(* IEC 61131-3 sources: s7-to-codesys/tests/POUs/ScenariosLang/FB_PumpInterlockLad_ScenarioTest, 6 files *)

(* ---- FB_PumpInterlockLad_ScenarioTest.decl.st ---- *)
// AUTO-GENERATED — не редактировать: s7conv gen-tests, сценарии scenarios/lang/FB_PumpInterlockLad.csv
// Правка — в CSV (scenarios/README.md), затем python -m s7conv build-corpus.
// Назначение: тесты поведения сконвертированного FB_PumpInterlockLad по сценариям CSV (сценариев: 5, строк: 25):
//             один метод-тест на сценарий, строки — по порядку с моделируемым временем GVL_S7Clock.
//             Ожидаемые значения — из CSV (эталонные модели по описанию логики блока), не из
//             результата конвертации.
// Автор:      s7conv 0.1.0 (сгенерировано)
// Версия:     не указана
// Документ:   scenarios/README.md, docs/methodology.md, раздел «Проверка поведения»
FUNCTION_BLOCK FB_PumpInterlockLad_ScenarioTest EXTENDS coUnit.FB_TestSuite
VAR
    fbAutoRunAndCount : FB_PumpInterlockLad;  // свой экземпляр на сценарий
    xAutoRunAndCountDone : BOOL;  // сценарий выполнен (выполняется один раз)
    fbLowLevelTripAndAck : FB_PumpInterlockLad;  // свой экземпляр на сценарий
    xLowLevelTripAndAckDone : BOOL;  // сценарий выполнен (выполняется один раз)
    fbHighPressure : FB_PumpInterlockLad;  // свой экземпляр на сценарий
    xHighPressureDone : BOOL;  // сценарий выполнен (выполняется один раз)
    fbMaintenanceJump : FB_PumpInterlockLad;  // свой экземпляр на сценарий
    xMaintenanceJumpDone : BOOL;  // сценарий выполнен (выполняется один раз)
    fbSetpointClamp : FB_PumpInterlockLad;  // свой экземпляр на сценарий
    xSetpointClampDone : BOOL;  // сценарий выполнен (выполняется один раз)
END_VAR

(* ---- AutoRunAndCount.method.impl.st ---- *)
// AUTO-GENERATED — не редактировать: scenarios/lang/FB_PumpInterlockLad.csv, сценарий AutoRunAndCount
coUnit.TEST('AutoRunAndCount');
IF NOT xAutoRunAndCountDone THEN
    xAutoRunAndCountDone := TRUE;
    GVL_S7Clock.xSimulation := TRUE;

    // #1, t = 0 мс — покой: уставка 0
    GVL_S7Clock.tSimNow := T#0MS;
    fbAutoRunAndCount.xAutoReq := FALSE;
    fbAutoRunAndCount.iLevel_cm := 120;
    fbAutoRunAndCount.iLevelMin_cm := 50;
    fbAutoRunAndCount.iPressure_kPa := 400;
    fbAutoRunAndCount.iPressureMax_kPa := 600;
    fbAutoRunAndCount.xAck := FALSE;
    fbAutoRunAndCount.xMaint := FALSE;
    fbAutoRunAndCount();
    AssertEquals_BOOL(Expected := FALSE, Actual := fbAutoRunAndCount.xPumpOn, Message := 'AutoRunAndCount#1 xPumpOn');
    AssertEquals_BOOL(Expected := FALSE,
                      Actual := fbAutoRunAndCount.xLowLevel,
                      Message := 'AutoRunAndCount#1 xLowLevel');
    AssertEquals_BOOL(Expected := FALSE,
                      Actual := fbAutoRunAndCount.xHighPress,
                      Message := 'AutoRunAndCount#1 xHighPress');
    AssertEquals_BOOL(Expected := FALSE, Actual := fbAutoRunAndCount.xAlarm, Message := 'AutoRunAndCount#1 xAlarm');
    AssertEquals_INT(Expected := 0, Actual := fbAutoRunAndCount.iRunCount, Message := 'AutoRunAndCount#1 iRunCount');
    AssertEquals_BOOL(Expected := FALSE, Actual := fbAutoRunAndCount.xCountOk, Message := 'AutoRunAndCount#1 xCountOk');
    AssertEquals_INT(Expected := 0,
                     Actual := fbAutoRunAndCount.iSetpoint_pct,
                     Message := 'AutoRunAndCount#1 iSetpoint_pct');
    AssertEquals_BOOL(Expected := FALSE, Actual := fbAutoRunAndCount.xChainOk, Message := 'AutoRunAndCount#1 xChainOk');
    AssertEquals_BOOL(Expected := FALSE, Actual := fbAutoRunAndCount.xRunMem, Message := 'AutoRunAndCount#1 xRunMem');

    // #2, t = 100 мс — включение №1: ENO = 1, уставка 120 → 100 → 90 → 80
    GVL_S7Clock.tSimNow := T#100MS;
    fbAutoRunAndCount.xAutoReq := TRUE;
    fbAutoRunAndCount();
    AssertEquals_BOOL(Expected := TRUE, Actual := fbAutoRunAndCount.xPumpOn, Message := 'AutoRunAndCount#2 xPumpOn');
    AssertEquals_BOOL(Expected := FALSE,
                      Actual := fbAutoRunAndCount.xLowLevel,
                      Message := 'AutoRunAndCount#2 xLowLevel');
    AssertEquals_BOOL(Expected := FALSE,
                      Actual := fbAutoRunAndCount.xHighPress,
                      Message := 'AutoRunAndCount#2 xHighPress');
    AssertEquals_BOOL(Expected := FALSE, Actual := fbAutoRunAndCount.xAlarm, Message := 'AutoRunAndCount#2 xAlarm');
    AssertEquals_INT(Expected := 1, Actual := fbAutoRunAndCount.iRunCount, Message := 'AutoRunAndCount#2 iRunCount');
    AssertEquals_BOOL(Expected := TRUE, Actual := fbAutoRunAndCount.xCountOk, Message := 'AutoRunAndCount#2 xCountOk');
    AssertEquals_INT(Expected := 80,
                     Actual := fbAutoRunAndCount.iSetpoint_pct,
                     Message := 'AutoRunAndCount#2 iSetpoint_pct');
    AssertEquals_BOOL(Expected := TRUE, Actual := fbAutoRunAndCount.xChainOk, Message := 'AutoRunAndCount#2 xChainOk');
    AssertEquals_BOOL(Expected := TRUE, Actual := fbAutoRunAndCount.xRunMem, Message := 'AutoRunAndCount#2 xRunMem');

    // #3, t = 200 мс — работает: фронта нет, ENO = 0
    GVL_S7Clock.tSimNow := T#200MS;
    fbAutoRunAndCount();
    AssertEquals_BOOL(Expected := TRUE, Actual := fbAutoRunAndCount.xPumpOn, Message := 'AutoRunAndCount#3 xPumpOn');
    AssertEquals_BOOL(Expected := FALSE,
                      Actual := fbAutoRunAndCount.xLowLevel,
                      Message := 'AutoRunAndCount#3 xLowLevel');
    AssertEquals_BOOL(Expected := FALSE,
                      Actual := fbAutoRunAndCount.xHighPress,
                      Message := 'AutoRunAndCount#3 xHighPress');
    AssertEquals_BOOL(Expected := FALSE, Actual := fbAutoRunAndCount.xAlarm, Message := 'AutoRunAndCount#3 xAlarm');
    AssertEquals_INT(Expected := 1, Actual := fbAutoRunAndCount.iRunCount, Message := 'AutoRunAndCount#3 iRunCount');
    AssertEquals_BOOL(Expected := FALSE, Actual := fbAutoRunAndCount.xCountOk, Message := 'AutoRunAndCount#3 xCountOk');
    AssertEquals_INT(Expected := 80,
                     Actual := fbAutoRunAndCount.iSetpoint_pct,
                     Message := 'AutoRunAndCount#3 iSetpoint_pct');
    AssertEquals_BOOL(Expected := TRUE, Actual := fbAutoRunAndCount.xChainOk, Message := 'AutoRunAndCount#3 xChainOk');
    AssertEquals_BOOL(Expected := TRUE, Actual := fbAutoRunAndCount.xRunMem, Message := 'AutoRunAndCount#3 xRunMem');

    // #4, t = 300 мс — запрос снят: насос выключен, уставка 0 (MOVE)
    GVL_S7Clock.tSimNow := T#300MS;
    fbAutoRunAndCount.xAutoReq := FALSE;
    fbAutoRunAndCount();
    AssertEquals_BOOL(Expected := FALSE, Actual := fbAutoRunAndCount.xPumpOn, Message := 'AutoRunAndCount#4 xPumpOn');
    AssertEquals_BOOL(Expected := FALSE,
                      Actual := fbAutoRunAndCount.xLowLevel,
                      Message := 'AutoRunAndCount#4 xLowLevel');
    AssertEquals_BOOL(Expected := FALSE,
                      Actual := fbAutoRunAndCount.xHighPress,
                      Message := 'AutoRunAndCount#4 xHighPress');
    AssertEquals_BOOL(Expected := FALSE, Actual := fbAutoRunAndCount.xAlarm, Message := 'AutoRunAndCount#4 xAlarm');
    AssertEquals_INT(Expected := 1, Actual := fbAutoRunAndCount.iRunCount, Message := 'AutoRunAndCount#4 iRunCount');
    AssertEquals_BOOL(Expected := FALSE, Actual := fbAutoRunAndCount.xCountOk, Message := 'AutoRunAndCount#4 xCountOk');
    AssertEquals_INT(Expected := 0,
                     Actual := fbAutoRunAndCount.iSetpoint_pct,
                     Message := 'AutoRunAndCount#4 iSetpoint_pct');
    AssertEquals_BOOL(Expected := FALSE, Actual := fbAutoRunAndCount.xChainOk, Message := 'AutoRunAndCount#4 xChainOk');
    AssertEquals_BOOL(Expected := FALSE, Actual := fbAutoRunAndCount.xRunMem, Message := 'AutoRunAndCount#4 xRunMem');

    // #5, t = 400 мс — включение №2
    GVL_S7Clock.tSimNow := T#400MS;
    fbAutoRunAndCount.xAutoReq := TRUE;
    fbAutoRunAndCount();
    AssertEquals_BOOL(Expected := TRUE, Actual := fbAutoRunAndCount.xPumpOn, Message := 'AutoRunAndCount#5 xPumpOn');
    AssertEquals_BOOL(Expected := FALSE,
                      Actual := fbAutoRunAndCount.xLowLevel,
                      Message := 'AutoRunAndCount#5 xLowLevel');
    AssertEquals_BOOL(Expected := FALSE,
                      Actual := fbAutoRunAndCount.xHighPress,
                      Message := 'AutoRunAndCount#5 xHighPress');
    AssertEquals_BOOL(Expected := FALSE, Actual := fbAutoRunAndCount.xAlarm, Message := 'AutoRunAndCount#5 xAlarm');
    AssertEquals_INT(Expected := 2, Actual := fbAutoRunAndCount.iRunCount, Message := 'AutoRunAndCount#5 iRunCount');
    AssertEquals_BOOL(Expected := TRUE, Actual := fbAutoRunAndCount.xCountOk, Message := 'AutoRunAndCount#5 xCountOk');
    AssertEquals_INT(Expected := 80,
                     Actual := fbAutoRunAndCount.iSetpoint_pct,
                     Message := 'AutoRunAndCount#5 iSetpoint_pct');
    AssertEquals_BOOL(Expected := TRUE, Actual := fbAutoRunAndCount.xChainOk, Message := 'AutoRunAndCount#5 xChainOk');
    AssertEquals_BOOL(Expected := TRUE, Actual := fbAutoRunAndCount.xRunMem, Message := 'AutoRunAndCount#5 xRunMem');

    GVL_S7Clock.xSimulation := FALSE;
END_IF
coUnit.TEST_FINISHED();

(* ---- HighPressure.method.impl.st ---- *)
// AUTO-GENERATED — не редактировать: scenarios/lang/FB_PumpInterlockLad.csv, сценарий HighPressure
coUnit.TEST('HighPressure');
IF NOT xHighPressureDone THEN
    xHighPressureDone := TRUE;
    GVL_S7Clock.xSimulation := TRUE;

    // #1, t = 0 мс — включение №1
    GVL_S7Clock.tSimNow := T#0MS;
    fbHighPressure.xAutoReq := TRUE;
    fbHighPressure.iLevel_cm := 120;
    fbHighPressure.iLevelMin_cm := 50;
    fbHighPressure.iPressure_kPa := 400;
    fbHighPressure.iPressureMax_kPa := 600;
    fbHighPressure.xAck := FALSE;
    fbHighPressure.xMaint := FALSE;
    fbHighPressure();
    AssertEquals_BOOL(Expected := TRUE, Actual := fbHighPressure.xPumpOn, Message := 'HighPressure#1 xPumpOn');
    AssertEquals_BOOL(Expected := FALSE, Actual := fbHighPressure.xLowLevel, Message := 'HighPressure#1 xLowLevel');
    AssertEquals_BOOL(Expected := FALSE, Actual := fbHighPressure.xHighPress, Message := 'HighPressure#1 xHighPress');
    AssertEquals_BOOL(Expected := FALSE, Actual := fbHighPressure.xAlarm, Message := 'HighPressure#1 xAlarm');
    AssertEquals_INT(Expected := 1, Actual := fbHighPressure.iRunCount, Message := 'HighPressure#1 iRunCount');
    AssertEquals_BOOL(Expected := TRUE, Actual := fbHighPressure.xCountOk, Message := 'HighPressure#1 xCountOk');
    AssertEquals_INT(Expected := 80, Actual := fbHighPressure.iSetpoint_pct, Message := 'HighPressure#1 iSetpoint_pct');
    AssertEquals_BOOL(Expected := TRUE, Actual := fbHighPressure.xChainOk, Message := 'HighPressure#1 xChainOk');
    AssertEquals_BOOL(Expected := TRUE, Actual := fbHighPressure.xRunMem, Message := 'HighPressure#1 xRunMem');

    // #2, t = 100 мс — 650 > 600: авария, насос выключен
    GVL_S7Clock.tSimNow := T#100MS;
    fbHighPressure.iPressure_kPa := 650;
    fbHighPressure();
    AssertEquals_BOOL(Expected := FALSE, Actual := fbHighPressure.xPumpOn, Message := 'HighPressure#2 xPumpOn');
    AssertEquals_BOOL(Expected := FALSE, Actual := fbHighPressure.xLowLevel, Message := 'HighPressure#2 xLowLevel');
    AssertEquals_BOOL(Expected := TRUE, Actual := fbHighPressure.xHighPress, Message := 'HighPressure#2 xHighPress');
    AssertEquals_BOOL(Expected := TRUE, Actual := fbHighPressure.xAlarm, Message := 'HighPressure#2 xAlarm');
    AssertEquals_INT(Expected := 1, Actual := fbHighPressure.iRunCount, Message := 'HighPressure#2 iRunCount');
    AssertEquals_BOOL(Expected := FALSE, Actual := fbHighPressure.xCountOk, Message := 'HighPressure#2 xCountOk');
    AssertEquals_INT(Expected := 0, Actual := fbHighPressure.iSetpoint_pct, Message := 'HighPressure#2 iSetpoint_pct');
    AssertEquals_BOOL(Expected := FALSE, Actual := fbHighPressure.xChainOk, Message := 'HighPressure#2 xChainOk');
    AssertEquals_BOOL(Expected := FALSE, Actual := fbHighPressure.xRunMem, Message := 'HighPressure#2 xRunMem');

    // #3, t = 200 мс — 600 не больше 600: квитирование снимает, включение №2
    GVL_S7Clock.tSimNow := T#200MS;
    fbHighPressure.iPressure_kPa := 600;
    fbHighPressure.xAck := TRUE;
    fbHighPressure();
    AssertEquals_BOOL(Expected := TRUE, Actual := fbHighPressure.xPumpOn, Message := 'HighPressure#3 xPumpOn');
    AssertEquals_BOOL(Expected := FALSE, Actual := fbHighPressure.xLowLevel, Message := 'HighPressure#3 xLowLevel');
    AssertEquals_BOOL(Expected := FALSE, Actual := fbHighPressure.xHighPress, Message := 'HighPressure#3 xHighPress');
    AssertEquals_BOOL(Expected := FALSE, Actual := fbHighPressure.xAlarm, Message := 'HighPressure#3 xAlarm');
    AssertEquals_INT(Expected := 2, Actual := fbHighPressure.iRunCount, Message := 'HighPressure#3 iRunCount');
    AssertEquals_BOOL(Expected := TRUE, Actual := fbHighPressure.xCountOk, Message := 'HighPressure#3 xCountOk');
    AssertEquals_INT(Expected := 80, Actual := fbHighPressure.iSetpoint_pct, Message := 'HighPressure#3 iSetpoint_pct');
    AssertEquals_BOOL(Expected := TRUE, Actual := fbHighPressure.xChainOk, Message := 'HighPressure#3 xChainOk');
    AssertEquals_BOOL(Expected := TRUE, Actual := fbHighPressure.xRunMem, Message := 'HighPressure#3 xRunMem');

    // #4, t = 300 мс — работает
    GVL_S7Clock.tSimNow := T#300MS;
    fbHighPressure.xAck := FALSE;
    fbHighPressure();
    AssertEquals_BOOL(Expected := TRUE, Actual := fbHighPressure.xPumpOn, Message := 'HighPressure#4 xPumpOn');
    AssertEquals_BOOL(Expected := FALSE, Actual := fbHighPressure.xLowLevel, Message := 'HighPressure#4 xLowLevel');
    AssertEquals_BOOL(Expected := FALSE, Actual := fbHighPressure.xHighPress, Message := 'HighPressure#4 xHighPress');
    AssertEquals_BOOL(Expected := FALSE, Actual := fbHighPressure.xAlarm, Message := 'HighPressure#4 xAlarm');
    AssertEquals_INT(Expected := 2, Actual := fbHighPressure.iRunCount, Message := 'HighPressure#4 iRunCount');
    AssertEquals_BOOL(Expected := FALSE, Actual := fbHighPressure.xCountOk, Message := 'HighPressure#4 xCountOk');
    AssertEquals_INT(Expected := 80, Actual := fbHighPressure.iSetpoint_pct, Message := 'HighPressure#4 iSetpoint_pct');
    AssertEquals_BOOL(Expected := TRUE, Actual := fbHighPressure.xChainOk, Message := 'HighPressure#4 xChainOk');
    AssertEquals_BOOL(Expected := TRUE, Actual := fbHighPressure.xRunMem, Message := 'HighPressure#4 xRunMem');

    GVL_S7Clock.xSimulation := FALSE;
END_IF
coUnit.TEST_FINISHED();

(* ---- LowLevelTripAndAck.method.impl.st ---- *)
// AUTO-GENERATED — не редактировать: scenarios/lang/FB_PumpInterlockLad.csv, сценарий LowLevelTripAndAck
coUnit.TEST('LowLevelTripAndAck');
IF NOT xLowLevelTripAndAckDone THEN
    xLowLevelTripAndAckDone := TRUE;
    GVL_S7Clock.xSimulation := TRUE;

    // #1, t = 0 мс — включение №1
    GVL_S7Clock.tSimNow := T#0MS;
    fbLowLevelTripAndAck.xAutoReq := TRUE;
    fbLowLevelTripAndAck.iLevel_cm := 120;
    fbLowLevelTripAndAck.iLevelMin_cm := 50;
    fbLowLevelTripAndAck.iPressure_kPa := 400;
    fbLowLevelTripAndAck.iPressureMax_kPa := 600;
    fbLowLevelTripAndAck.xAck := FALSE;
    fbLowLevelTripAndAck.xMaint := FALSE;
    fbLowLevelTripAndAck();
    AssertEquals_BOOL(Expected := TRUE,
                      Actual := fbLowLevelTripAndAck.xPumpOn,
                      Message := 'LowLevelTripAndAck#1 xPumpOn');
    AssertEquals_BOOL(Expected := FALSE,
                      Actual := fbLowLevelTripAndAck.xLowLevel,
                      Message := 'LowLevelTripAndAck#1 xLowLevel');
    AssertEquals_BOOL(Expected := FALSE,
                      Actual := fbLowLevelTripAndAck.xHighPress,
                      Message := 'LowLevelTripAndAck#1 xHighPress');
    AssertEquals_BOOL(Expected := FALSE,
                      Actual := fbLowLevelTripAndAck.xAlarm,
                      Message := 'LowLevelTripAndAck#1 xAlarm');
    AssertEquals_INT(Expected := 1,
                     Actual := fbLowLevelTripAndAck.iRunCount,
                     Message := 'LowLevelTripAndAck#1 iRunCount');
    AssertEquals_BOOL(Expected := TRUE,
                      Actual := fbLowLevelTripAndAck.xCountOk,
                      Message := 'LowLevelTripAndAck#1 xCountOk');
    AssertEquals_INT(Expected := 80,
                     Actual := fbLowLevelTripAndAck.iSetpoint_pct,
                     Message := 'LowLevelTripAndAck#1 iSetpoint_pct');
    AssertEquals_BOOL(Expected := TRUE,
                      Actual := fbLowLevelTripAndAck.xChainOk,
                      Message := 'LowLevelTripAndAck#1 xChainOk');
    AssertEquals_BOOL(Expected := TRUE,
                      Actual := fbLowLevelTripAndAck.xRunMem,
                      Message := 'LowLevelTripAndAck#1 xRunMem');

    // #2, t = 100 мс — уровень 40 < 50: авария, насос выключен
    GVL_S7Clock.tSimNow := T#100MS;
    fbLowLevelTripAndAck.iLevel_cm := 40;
    fbLowLevelTripAndAck();
    AssertEquals_BOOL(Expected := FALSE,
                      Actual := fbLowLevelTripAndAck.xPumpOn,
                      Message := 'LowLevelTripAndAck#2 xPumpOn');
    AssertEquals_BOOL(Expected := TRUE,
                      Actual := fbLowLevelTripAndAck.xLowLevel,
                      Message := 'LowLevelTripAndAck#2 xLowLevel');
    AssertEquals_BOOL(Expected := FALSE,
                      Actual := fbLowLevelTripAndAck.xHighPress,
                      Message := 'LowLevelTripAndAck#2 xHighPress');
    AssertEquals_BOOL(Expected := TRUE,
                      Actual := fbLowLevelTripAndAck.xAlarm,
                      Message := 'LowLevelTripAndAck#2 xAlarm');
    AssertEquals_INT(Expected := 1,
                     Actual := fbLowLevelTripAndAck.iRunCount,
                     Message := 'LowLevelTripAndAck#2 iRunCount');
    AssertEquals_BOOL(Expected := FALSE,
                      Actual := fbLowLevelTripAndAck.xCountOk,
                      Message := 'LowLevelTripAndAck#2 xCountOk');
    AssertEquals_INT(Expected := 0,
                     Actual := fbLowLevelTripAndAck.iSetpoint_pct,
                     Message := 'LowLevelTripAndAck#2 iSetpoint_pct');
    AssertEquals_BOOL(Expected := FALSE,
                      Actual := fbLowLevelTripAndAck.xChainOk,
                      Message := 'LowLevelTripAndAck#2 xChainOk');
    AssertEquals_BOOL(Expected := FALSE,
                      Actual := fbLowLevelTripAndAck.xRunMem,
                      Message := 'LowLevelTripAndAck#2 xRunMem');

    // #3, t = 200 мс — уровень в норме: авария держится
    GVL_S7Clock.tSimNow := T#200MS;
    fbLowLevelTripAndAck.iLevel_cm := 60;
    fbLowLevelTripAndAck();
    AssertEquals_BOOL(Expected := FALSE,
                      Actual := fbLowLevelTripAndAck.xPumpOn,
                      Message := 'LowLevelTripAndAck#3 xPumpOn');
    AssertEquals_BOOL(Expected := FALSE,
                      Actual := fbLowLevelTripAndAck.xLowLevel,
                      Message := 'LowLevelTripAndAck#3 xLowLevel');
    AssertEquals_BOOL(Expected := FALSE,
                      Actual := fbLowLevelTripAndAck.xHighPress,
                      Message := 'LowLevelTripAndAck#3 xHighPress');
    AssertEquals_BOOL(Expected := TRUE,
                      Actual := fbLowLevelTripAndAck.xAlarm,
                      Message := 'LowLevelTripAndAck#3 xAlarm');
    AssertEquals_INT(Expected := 1,
                     Actual := fbLowLevelTripAndAck.iRunCount,
                     Message := 'LowLevelTripAndAck#3 iRunCount');
    AssertEquals_BOOL(Expected := FALSE,
                      Actual := fbLowLevelTripAndAck.xCountOk,
                      Message := 'LowLevelTripAndAck#3 xCountOk');
    AssertEquals_INT(Expected := 0,
                     Actual := fbLowLevelTripAndAck.iSetpoint_pct,
                     Message := 'LowLevelTripAndAck#3 iSetpoint_pct');
    AssertEquals_BOOL(Expected := FALSE,
                      Actual := fbLowLevelTripAndAck.xChainOk,
                      Message := 'LowLevelTripAndAck#3 xChainOk');
    AssertEquals_BOOL(Expected := FALSE,
                      Actual := fbLowLevelTripAndAck.xRunMem,
                      Message := 'LowLevelTripAndAck#3 xRunMem');

    // #4, t = 300 мс — квитирование при низком уровне: не снимается
    GVL_S7Clock.tSimNow := T#300MS;
    fbLowLevelTripAndAck.iLevel_cm := 45;
    fbLowLevelTripAndAck.xAck := TRUE;
    fbLowLevelTripAndAck();
    AssertEquals_BOOL(Expected := FALSE,
                      Actual := fbLowLevelTripAndAck.xPumpOn,
                      Message := 'LowLevelTripAndAck#4 xPumpOn');
    AssertEquals_BOOL(Expected := TRUE,
                      Actual := fbLowLevelTripAndAck.xLowLevel,
                      Message := 'LowLevelTripAndAck#4 xLowLevel');
    AssertEquals_BOOL(Expected := FALSE,
                      Actual := fbLowLevelTripAndAck.xHighPress,
                      Message := 'LowLevelTripAndAck#4 xHighPress');
    AssertEquals_BOOL(Expected := TRUE,
                      Actual := fbLowLevelTripAndAck.xAlarm,
                      Message := 'LowLevelTripAndAck#4 xAlarm');
    AssertEquals_INT(Expected := 1,
                     Actual := fbLowLevelTripAndAck.iRunCount,
                     Message := 'LowLevelTripAndAck#4 iRunCount');
    AssertEquals_BOOL(Expected := FALSE,
                      Actual := fbLowLevelTripAndAck.xCountOk,
                      Message := 'LowLevelTripAndAck#4 xCountOk');
    AssertEquals_INT(Expected := 0,
                     Actual := fbLowLevelTripAndAck.iSetpoint_pct,
                     Message := 'LowLevelTripAndAck#4 iSetpoint_pct');
    AssertEquals_BOOL(Expected := FALSE,
                      Actual := fbLowLevelTripAndAck.xChainOk,
                      Message := 'LowLevelTripAndAck#4 xChainOk');
    AssertEquals_BOOL(Expected := FALSE,
                      Actual := fbLowLevelTripAndAck.xRunMem,
                      Message := 'LowLevelTripAndAck#4 xRunMem');

    // #5, t = 400 мс — уровень в норме при нажатом квитировании: снята, включение №2
    GVL_S7Clock.tSimNow := T#400MS;
    fbLowLevelTripAndAck.iLevel_cm := 70;
    fbLowLevelTripAndAck();
    AssertEquals_BOOL(Expected := TRUE,
                      Actual := fbLowLevelTripAndAck.xPumpOn,
                      Message := 'LowLevelTripAndAck#5 xPumpOn');
    AssertEquals_BOOL(Expected := FALSE,
                      Actual := fbLowLevelTripAndAck.xLowLevel,
                      Message := 'LowLevelTripAndAck#5 xLowLevel');
    AssertEquals_BOOL(Expected := FALSE,
                      Actual := fbLowLevelTripAndAck.xHighPress,
                      Message := 'LowLevelTripAndAck#5 xHighPress');
    AssertEquals_BOOL(Expected := FALSE,
                      Actual := fbLowLevelTripAndAck.xAlarm,
                      Message := 'LowLevelTripAndAck#5 xAlarm');
    AssertEquals_INT(Expected := 2,
                     Actual := fbLowLevelTripAndAck.iRunCount,
                     Message := 'LowLevelTripAndAck#5 iRunCount');
    AssertEquals_BOOL(Expected := TRUE,
                      Actual := fbLowLevelTripAndAck.xCountOk,
                      Message := 'LowLevelTripAndAck#5 xCountOk');
    AssertEquals_INT(Expected := 70,
                     Actual := fbLowLevelTripAndAck.iSetpoint_pct,
                     Message := 'LowLevelTripAndAck#5 iSetpoint_pct');
    AssertEquals_BOOL(Expected := TRUE,
                      Actual := fbLowLevelTripAndAck.xChainOk,
                      Message := 'LowLevelTripAndAck#5 xChainOk');
    AssertEquals_BOOL(Expected := TRUE,
                      Actual := fbLowLevelTripAndAck.xRunMem,
                      Message := 'LowLevelTripAndAck#5 xRunMem');

    // #6, t = 500 мс — работает
    GVL_S7Clock.tSimNow := T#500MS;
    fbLowLevelTripAndAck.xAck := FALSE;
    fbLowLevelTripAndAck();
    AssertEquals_BOOL(Expected := TRUE,
                      Actual := fbLowLevelTripAndAck.xPumpOn,
                      Message := 'LowLevelTripAndAck#6 xPumpOn');
    AssertEquals_BOOL(Expected := FALSE,
                      Actual := fbLowLevelTripAndAck.xLowLevel,
                      Message := 'LowLevelTripAndAck#6 xLowLevel');
    AssertEquals_BOOL(Expected := FALSE,
                      Actual := fbLowLevelTripAndAck.xHighPress,
                      Message := 'LowLevelTripAndAck#6 xHighPress');
    AssertEquals_BOOL(Expected := FALSE,
                      Actual := fbLowLevelTripAndAck.xAlarm,
                      Message := 'LowLevelTripAndAck#6 xAlarm');
    AssertEquals_INT(Expected := 2,
                     Actual := fbLowLevelTripAndAck.iRunCount,
                     Message := 'LowLevelTripAndAck#6 iRunCount');
    AssertEquals_BOOL(Expected := FALSE,
                      Actual := fbLowLevelTripAndAck.xCountOk,
                      Message := 'LowLevelTripAndAck#6 xCountOk');
    AssertEquals_INT(Expected := 70,
                     Actual := fbLowLevelTripAndAck.iSetpoint_pct,
                     Message := 'LowLevelTripAndAck#6 iSetpoint_pct');
    AssertEquals_BOOL(Expected := TRUE,
                      Actual := fbLowLevelTripAndAck.xChainOk,
                      Message := 'LowLevelTripAndAck#6 xChainOk');
    AssertEquals_BOOL(Expected := TRUE,
                      Actual := fbLowLevelTripAndAck.xRunMem,
                      Message := 'LowLevelTripAndAck#6 xRunMem');

    GVL_S7Clock.xSimulation := FALSE;
END_IF
coUnit.TEST_FINISHED();

(* ---- MaintenanceJump.method.impl.st ---- *)
// AUTO-GENERATED — не редактировать: scenarios/lang/FB_PumpInterlockLad.csv, сценарий MaintenanceJump
coUnit.TEST('MaintenanceJump');
IF NOT xMaintenanceJumpDone THEN
    xMaintenanceJumpDone := TRUE;
    GVL_S7Clock.xSimulation := TRUE;

    // #1, t = 0 мс — включение №1, xCountOk = 1
    GVL_S7Clock.tSimNow := T#0MS;
    fbMaintenanceJump.xAutoReq := TRUE;
    fbMaintenanceJump.iLevel_cm := 120;
    fbMaintenanceJump.iLevelMin_cm := 50;
    fbMaintenanceJump.iPressure_kPa := 400;
    fbMaintenanceJump.iPressureMax_kPa := 600;
    fbMaintenanceJump.xAck := FALSE;
    fbMaintenanceJump.xMaint := FALSE;
    fbMaintenanceJump();
    AssertEquals_BOOL(Expected := TRUE, Actual := fbMaintenanceJump.xPumpOn, Message := 'MaintenanceJump#1 xPumpOn');
    AssertEquals_BOOL(Expected := FALSE,
                      Actual := fbMaintenanceJump.xLowLevel,
                      Message := 'MaintenanceJump#1 xLowLevel');
    AssertEquals_BOOL(Expected := FALSE,
                      Actual := fbMaintenanceJump.xHighPress,
                      Message := 'MaintenanceJump#1 xHighPress');
    AssertEquals_BOOL(Expected := FALSE, Actual := fbMaintenanceJump.xAlarm, Message := 'MaintenanceJump#1 xAlarm');
    AssertEquals_INT(Expected := 1, Actual := fbMaintenanceJump.iRunCount, Message := 'MaintenanceJump#1 iRunCount');
    AssertEquals_BOOL(Expected := TRUE, Actual := fbMaintenanceJump.xCountOk, Message := 'MaintenanceJump#1 xCountOk');
    AssertEquals_INT(Expected := 80,
                     Actual := fbMaintenanceJump.iSetpoint_pct,
                     Message := 'MaintenanceJump#1 iSetpoint_pct');
    AssertEquals_BOOL(Expected := TRUE, Actual := fbMaintenanceJump.xChainOk, Message := 'MaintenanceJump#1 xChainOk');
    AssertEquals_BOOL(Expected := TRUE, Actual := fbMaintenanceJump.xRunMem, Message := 'MaintenanceJump#1 xRunMem');

    // #2, t = 100 мс — обслуживание: насос выключен; xCountOk и xRunMem сохраняют значения
    GVL_S7Clock.tSimNow := T#100MS;
    fbMaintenanceJump.xMaint := TRUE;
    fbMaintenanceJump();
    AssertEquals_BOOL(Expected := FALSE, Actual := fbMaintenanceJump.xPumpOn, Message := 'MaintenanceJump#2 xPumpOn');
    AssertEquals_BOOL(Expected := FALSE,
                      Actual := fbMaintenanceJump.xLowLevel,
                      Message := 'MaintenanceJump#2 xLowLevel');
    AssertEquals_BOOL(Expected := FALSE,
                      Actual := fbMaintenanceJump.xHighPress,
                      Message := 'MaintenanceJump#2 xHighPress');
    AssertEquals_BOOL(Expected := FALSE, Actual := fbMaintenanceJump.xAlarm, Message := 'MaintenanceJump#2 xAlarm');
    AssertEquals_INT(Expected := 1, Actual := fbMaintenanceJump.iRunCount, Message := 'MaintenanceJump#2 iRunCount');
    AssertEquals_BOOL(Expected := TRUE, Actual := fbMaintenanceJump.xCountOk, Message := 'MaintenanceJump#2 xCountOk');
    AssertEquals_INT(Expected := 0,
                     Actual := fbMaintenanceJump.iSetpoint_pct,
                     Message := 'MaintenanceJump#2 iSetpoint_pct');
    AssertEquals_BOOL(Expected := FALSE, Actual := fbMaintenanceJump.xChainOk, Message := 'MaintenanceJump#2 xChainOk');
    AssertEquals_BOOL(Expected := TRUE, Actual := fbMaintenanceJump.xRunMem, Message := 'MaintenanceJump#2 xRunMem');

    // #3, t = 200 мс — обслуживание держится
    GVL_S7Clock.tSimNow := T#200MS;
    fbMaintenanceJump();
    AssertEquals_BOOL(Expected := FALSE, Actual := fbMaintenanceJump.xPumpOn, Message := 'MaintenanceJump#3 xPumpOn');
    AssertEquals_BOOL(Expected := FALSE,
                      Actual := fbMaintenanceJump.xLowLevel,
                      Message := 'MaintenanceJump#3 xLowLevel');
    AssertEquals_BOOL(Expected := FALSE,
                      Actual := fbMaintenanceJump.xHighPress,
                      Message := 'MaintenanceJump#3 xHighPress');
    AssertEquals_BOOL(Expected := FALSE, Actual := fbMaintenanceJump.xAlarm, Message := 'MaintenanceJump#3 xAlarm');
    AssertEquals_INT(Expected := 1, Actual := fbMaintenanceJump.iRunCount, Message := 'MaintenanceJump#3 iRunCount');
    AssertEquals_BOOL(Expected := TRUE, Actual := fbMaintenanceJump.xCountOk, Message := 'MaintenanceJump#3 xCountOk');
    AssertEquals_INT(Expected := 0,
                     Actual := fbMaintenanceJump.iSetpoint_pct,
                     Message := 'MaintenanceJump#3 iSetpoint_pct');
    AssertEquals_BOOL(Expected := FALSE, Actual := fbMaintenanceJump.xChainOk, Message := 'MaintenanceJump#3 xChainOk');
    AssertEquals_BOOL(Expected := TRUE, Actual := fbMaintenanceJump.xRunMem, Message := 'MaintenanceJump#3 xRunMem');

    // #4, t = 300 мс — выход из обслуживания: насос включён, фронта нет — бит памяти остался 1
    GVL_S7Clock.tSimNow := T#300MS;
    fbMaintenanceJump.xMaint := FALSE;
    fbMaintenanceJump();
    AssertEquals_BOOL(Expected := TRUE, Actual := fbMaintenanceJump.xPumpOn, Message := 'MaintenanceJump#4 xPumpOn');
    AssertEquals_BOOL(Expected := FALSE,
                      Actual := fbMaintenanceJump.xLowLevel,
                      Message := 'MaintenanceJump#4 xLowLevel');
    AssertEquals_BOOL(Expected := FALSE,
                      Actual := fbMaintenanceJump.xHighPress,
                      Message := 'MaintenanceJump#4 xHighPress');
    AssertEquals_BOOL(Expected := FALSE, Actual := fbMaintenanceJump.xAlarm, Message := 'MaintenanceJump#4 xAlarm');
    AssertEquals_INT(Expected := 1, Actual := fbMaintenanceJump.iRunCount, Message := 'MaintenanceJump#4 iRunCount');
    AssertEquals_BOOL(Expected := FALSE, Actual := fbMaintenanceJump.xCountOk, Message := 'MaintenanceJump#4 xCountOk');
    AssertEquals_INT(Expected := 80,
                     Actual := fbMaintenanceJump.iSetpoint_pct,
                     Message := 'MaintenanceJump#4 iSetpoint_pct');
    AssertEquals_BOOL(Expected := TRUE, Actual := fbMaintenanceJump.xChainOk, Message := 'MaintenanceJump#4 xChainOk');
    AssertEquals_BOOL(Expected := TRUE, Actual := fbMaintenanceJump.xRunMem, Message := 'MaintenanceJump#4 xRunMem');

    // #5, t = 400 мс — запрос снят
    GVL_S7Clock.tSimNow := T#400MS;
    fbMaintenanceJump.xAutoReq := FALSE;
    fbMaintenanceJump();
    AssertEquals_BOOL(Expected := FALSE, Actual := fbMaintenanceJump.xPumpOn, Message := 'MaintenanceJump#5 xPumpOn');
    AssertEquals_BOOL(Expected := FALSE,
                      Actual := fbMaintenanceJump.xLowLevel,
                      Message := 'MaintenanceJump#5 xLowLevel');
    AssertEquals_BOOL(Expected := FALSE,
                      Actual := fbMaintenanceJump.xHighPress,
                      Message := 'MaintenanceJump#5 xHighPress');
    AssertEquals_BOOL(Expected := FALSE, Actual := fbMaintenanceJump.xAlarm, Message := 'MaintenanceJump#5 xAlarm');
    AssertEquals_INT(Expected := 1, Actual := fbMaintenanceJump.iRunCount, Message := 'MaintenanceJump#5 iRunCount');
    AssertEquals_BOOL(Expected := FALSE, Actual := fbMaintenanceJump.xCountOk, Message := 'MaintenanceJump#5 xCountOk');
    AssertEquals_INT(Expected := 0,
                     Actual := fbMaintenanceJump.iSetpoint_pct,
                     Message := 'MaintenanceJump#5 iSetpoint_pct');
    AssertEquals_BOOL(Expected := FALSE, Actual := fbMaintenanceJump.xChainOk, Message := 'MaintenanceJump#5 xChainOk');
    AssertEquals_BOOL(Expected := FALSE, Actual := fbMaintenanceJump.xRunMem, Message := 'MaintenanceJump#5 xRunMem');

    // #6, t = 500 мс — включение №2
    GVL_S7Clock.tSimNow := T#500MS;
    fbMaintenanceJump.xAutoReq := TRUE;
    fbMaintenanceJump();
    AssertEquals_BOOL(Expected := TRUE, Actual := fbMaintenanceJump.xPumpOn, Message := 'MaintenanceJump#6 xPumpOn');
    AssertEquals_BOOL(Expected := FALSE,
                      Actual := fbMaintenanceJump.xLowLevel,
                      Message := 'MaintenanceJump#6 xLowLevel');
    AssertEquals_BOOL(Expected := FALSE,
                      Actual := fbMaintenanceJump.xHighPress,
                      Message := 'MaintenanceJump#6 xHighPress');
    AssertEquals_BOOL(Expected := FALSE, Actual := fbMaintenanceJump.xAlarm, Message := 'MaintenanceJump#6 xAlarm');
    AssertEquals_INT(Expected := 2, Actual := fbMaintenanceJump.iRunCount, Message := 'MaintenanceJump#6 iRunCount');
    AssertEquals_BOOL(Expected := TRUE, Actual := fbMaintenanceJump.xCountOk, Message := 'MaintenanceJump#6 xCountOk');
    AssertEquals_INT(Expected := 80,
                     Actual := fbMaintenanceJump.iSetpoint_pct,
                     Message := 'MaintenanceJump#6 iSetpoint_pct');
    AssertEquals_BOOL(Expected := TRUE, Actual := fbMaintenanceJump.xChainOk, Message := 'MaintenanceJump#6 xChainOk');
    AssertEquals_BOOL(Expected := TRUE, Actual := fbMaintenanceJump.xRunMem, Message := 'MaintenanceJump#6 xRunMem');

    GVL_S7Clock.xSimulation := FALSE;
END_IF
coUnit.TEST_FINISHED();

(* ---- SetpointClamp.method.impl.st ---- *)
// AUTO-GENERATED — не редактировать: scenarios/lang/FB_PumpInterlockLad.csv, сценарий SetpointClamp
coUnit.TEST('SetpointClamp');
IF NOT xSetpointClampDone THEN
    xSetpointClampDone := TRUE;
    GVL_S7Clock.xSimulation := TRUE;

    // #1, t = 0 мс — 55 → 55 → 55 → 55
    GVL_S7Clock.tSimNow := T#0MS;
    fbSetpointClamp.xAutoReq := TRUE;
    fbSetpointClamp.iLevel_cm := 55;
    fbSetpointClamp.iLevelMin_cm := 50;
    fbSetpointClamp.iPressure_kPa := 400;
    fbSetpointClamp.iPressureMax_kPa := 600;
    fbSetpointClamp.xAck := FALSE;
    fbSetpointClamp.xMaint := FALSE;
    fbSetpointClamp();
    AssertEquals_BOOL(Expected := TRUE, Actual := fbSetpointClamp.xPumpOn, Message := 'SetpointClamp#1 xPumpOn');
    AssertEquals_BOOL(Expected := FALSE, Actual := fbSetpointClamp.xLowLevel, Message := 'SetpointClamp#1 xLowLevel');
    AssertEquals_BOOL(Expected := FALSE, Actual := fbSetpointClamp.xHighPress, Message := 'SetpointClamp#1 xHighPress');
    AssertEquals_BOOL(Expected := FALSE, Actual := fbSetpointClamp.xAlarm, Message := 'SetpointClamp#1 xAlarm');
    AssertEquals_INT(Expected := 1, Actual := fbSetpointClamp.iRunCount, Message := 'SetpointClamp#1 iRunCount');
    AssertEquals_BOOL(Expected := TRUE, Actual := fbSetpointClamp.xCountOk, Message := 'SetpointClamp#1 xCountOk');
    AssertEquals_INT(Expected := 55,
                     Actual := fbSetpointClamp.iSetpoint_pct,
                     Message := 'SetpointClamp#1 iSetpoint_pct');
    AssertEquals_BOOL(Expected := TRUE, Actual := fbSetpointClamp.xChainOk, Message := 'SetpointClamp#1 xChainOk');
    AssertEquals_BOOL(Expected := TRUE, Actual := fbSetpointClamp.xRunMem, Message := 'SetpointClamp#1 xRunMem');

    // #2, t = 100 мс — 95 → 95 → 90 → 80
    GVL_S7Clock.tSimNow := T#100MS;
    fbSetpointClamp.iLevel_cm := 95;
    fbSetpointClamp();
    AssertEquals_BOOL(Expected := TRUE, Actual := fbSetpointClamp.xPumpOn, Message := 'SetpointClamp#2 xPumpOn');
    AssertEquals_BOOL(Expected := FALSE, Actual := fbSetpointClamp.xLowLevel, Message := 'SetpointClamp#2 xLowLevel');
    AssertEquals_BOOL(Expected := FALSE, Actual := fbSetpointClamp.xHighPress, Message := 'SetpointClamp#2 xHighPress');
    AssertEquals_BOOL(Expected := FALSE, Actual := fbSetpointClamp.xAlarm, Message := 'SetpointClamp#2 xAlarm');
    AssertEquals_INT(Expected := 1, Actual := fbSetpointClamp.iRunCount, Message := 'SetpointClamp#2 iRunCount');
    AssertEquals_BOOL(Expected := FALSE, Actual := fbSetpointClamp.xCountOk, Message := 'SetpointClamp#2 xCountOk');
    AssertEquals_INT(Expected := 80,
                     Actual := fbSetpointClamp.iSetpoint_pct,
                     Message := 'SetpointClamp#2 iSetpoint_pct');
    AssertEquals_BOOL(Expected := TRUE, Actual := fbSetpointClamp.xChainOk, Message := 'SetpointClamp#2 xChainOk');
    AssertEquals_BOOL(Expected := TRUE, Actual := fbSetpointClamp.xRunMem, Message := 'SetpointClamp#2 xRunMem');

    // #3, t = 200 мс — 15 → 15 → 15 → 20
    GVL_S7Clock.tSimNow := T#200MS;
    fbSetpointClamp.iLevel_cm := 15;
    fbSetpointClamp.iLevelMin_cm := 10;
    fbSetpointClamp();
    AssertEquals_BOOL(Expected := TRUE, Actual := fbSetpointClamp.xPumpOn, Message := 'SetpointClamp#3 xPumpOn');
    AssertEquals_BOOL(Expected := FALSE, Actual := fbSetpointClamp.xLowLevel, Message := 'SetpointClamp#3 xLowLevel');
    AssertEquals_BOOL(Expected := FALSE, Actual := fbSetpointClamp.xHighPress, Message := 'SetpointClamp#3 xHighPress');
    AssertEquals_BOOL(Expected := FALSE, Actual := fbSetpointClamp.xAlarm, Message := 'SetpointClamp#3 xAlarm');
    AssertEquals_INT(Expected := 1, Actual := fbSetpointClamp.iRunCount, Message := 'SetpointClamp#3 iRunCount');
    AssertEquals_BOOL(Expected := FALSE, Actual := fbSetpointClamp.xCountOk, Message := 'SetpointClamp#3 xCountOk');
    AssertEquals_INT(Expected := 20,
                     Actual := fbSetpointClamp.iSetpoint_pct,
                     Message := 'SetpointClamp#3 iSetpoint_pct');
    AssertEquals_BOOL(Expected := TRUE, Actual := fbSetpointClamp.xChainOk, Message := 'SetpointClamp#3 xChainOk');
    AssertEquals_BOOL(Expected := TRUE, Actual := fbSetpointClamp.xRunMem, Message := 'SetpointClamp#3 xRunMem');

    // #4, t = 300 мс — 5 → 5 → 10 → 20
    GVL_S7Clock.tSimNow := T#300MS;
    fbSetpointClamp.iLevel_cm := 5;
    fbSetpointClamp.iLevelMin_cm := 0;
    fbSetpointClamp();
    AssertEquals_BOOL(Expected := TRUE, Actual := fbSetpointClamp.xPumpOn, Message := 'SetpointClamp#4 xPumpOn');
    AssertEquals_BOOL(Expected := FALSE, Actual := fbSetpointClamp.xLowLevel, Message := 'SetpointClamp#4 xLowLevel');
    AssertEquals_BOOL(Expected := FALSE, Actual := fbSetpointClamp.xHighPress, Message := 'SetpointClamp#4 xHighPress');
    AssertEquals_BOOL(Expected := FALSE, Actual := fbSetpointClamp.xAlarm, Message := 'SetpointClamp#4 xAlarm');
    AssertEquals_INT(Expected := 1, Actual := fbSetpointClamp.iRunCount, Message := 'SetpointClamp#4 iRunCount');
    AssertEquals_BOOL(Expected := FALSE, Actual := fbSetpointClamp.xCountOk, Message := 'SetpointClamp#4 xCountOk');
    AssertEquals_INT(Expected := 20,
                     Actual := fbSetpointClamp.iSetpoint_pct,
                     Message := 'SetpointClamp#4 iSetpoint_pct');
    AssertEquals_BOOL(Expected := TRUE, Actual := fbSetpointClamp.xChainOk, Message := 'SetpointClamp#4 xChainOk');
    AssertEquals_BOOL(Expected := TRUE, Actual := fbSetpointClamp.xRunMem, Message := 'SetpointClamp#4 xRunMem');

    GVL_S7Clock.xSimulation := FALSE;
END_IF
coUnit.TEST_FINISHED();
